// TIA Portal V21 export
// export: Created 2026-11-11T00:47:54.2994255Z, ExportSetting WithDefaults, DisplayName Totally Integrated Automation Portal, DisplayVersion V21 Update 3, DisplayName STEP 7 Professional, DisplayVersion V21 Update 3, DisplayName STEP 7 Safety, DisplayVersion V21, DisplayName Tech WebApplication, DisplayVersion V21, DisplayName WinCC Basic/Comfort/Advanced, DisplayVersion V21 Update 3, DisplayName WinCC Unified, DisplayVersion V21 Update 3
FUNCTION_BLOCK "FB_Lad_ex122"   // FB397, LAD
{ S7_Optimized_Access := 'TRUE' }
VERSION : 0.1
// stored: AutoNumber true, IsIECCheckEnabled false, IsRetainMemResEnabled false, MemoryReserve 100, SetENOAutomatically false, UDAEnableTagReadback false
   VAR_INPUT
      v_operatemode : Byte;
      v_datamode : Byte;
      v_dispclassnr : Array[0..31] of UInt;
      v_lcid : UDInt;
   END_VAR
   VAR_OUTPUT
      v_dataready : Bool;
      v_busy : Bool;
      v_error : Bool;
      v_init : Bool;
      v_status : Word;
   END_VAR
   VAR_IN_OUT
      v_data : AlarmData;
   END_VAR
   VAR
      inst { S7_SetPoint := 'True'} : Get_Alarm;
   END_VAR
BEGIN

REGION Network 1: Get_Alarm - Read pending alarm
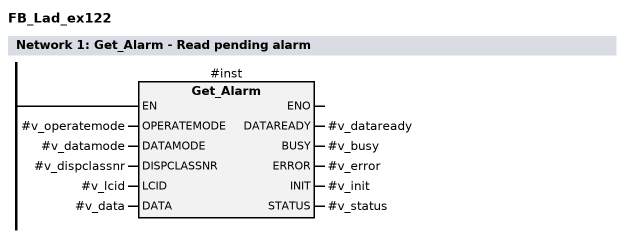
   RUNG wire#powerrail
      #inst.Get_Alarm(OperateMode := #v_operatemode, DataMode := #v_datamode, DispClassNr := #v_dispclassnr, Lcid := #v_lcid, Data := #v_data, DataReady => #v_dataready, Busy => #v_busy, Error => #v_error, Init => #v_init, Status => #v_status)
   END_RUNG
   // the same network as SCL:
   #inst(OperateMode := #v_operatemode,   // Get_Alarm
         DataMode := #v_datamode,
         DispClassNr := #v_dispclassnr,
         Lcid := #v_lcid,
         Data := #v_data,
         DataReady => #v_dataready,
         Busy => #v_busy,
         Error => #v_error,
         Init => #v_init,
         Status => #v_status);
END_REGION
END_FUNCTION_BLOCK
